FUNCTION_BLOCK "Tgp_CTU_LimitDriver_LAD"
{ S7_Optimized_Access := 'TRUE' }
VAR_INPUT
    Edges : Int;
    Reset : Bool;
END_VAR
VAR_OUTPUT
    Count : Int;
    Done : Bool;
    Rejected : Bool;
END_VAR
VAR
    // COUNTER is a reserved SCL data type keyword, so the instance has a distinct name.
    CtuInstance : "Tgp_CTU_LAD";
END_VAR
VAR_TEMP
    Index : Int;
END_VAR
BEGIN
    #Rejected := (#Edges < 0) OR (#Edges > 512);
    IF NOT #Rejected THEN
        IF #Reset OR (#Edges = 0) THEN
            #CtuInstance(Enable := FALSE, Down := FALSE, Reset := #Reset,
                     Load := FALSE, Preset := 32767,
                     Done => #Done, Count => #Count);
        ELSE
            FOR #Index := 1 TO #Edges DO
                #CtuInstance(Enable := FALSE, Down := FALSE, Reset := FALSE,
                         Load := FALSE, Preset := 32767,
                         Done => #Done, Count => #Count);
                #CtuInstance(Enable := TRUE, Down := FALSE, Reset := FALSE,
                         Load := FALSE, Preset := 32767,
                         Done => #Done, Count => #Count);
            END_FOR;
        END_IF;
    END_IF;
END_FUNCTION_BLOCK
